{attribute 'qualified_only'}
VAR_GLOBAL
    // Failure hooks for the simulated devices, set from the HMI or a watch
    // window. Each one acts only while its device is simulated.
    TankValveStuck  : BOOL;
    DrainValveStuck : BOOL;
    LiftStuck       : BOOL;
    SlideStuck      : BOOL;
    GripperStuck    : BOOL;
END_VAR

(* stored: Version 1.1.0.1
   GVL GVL_Sim: Id {afc57dfd-7eaf-4cce-aeb0-6919f986cd06} *)
